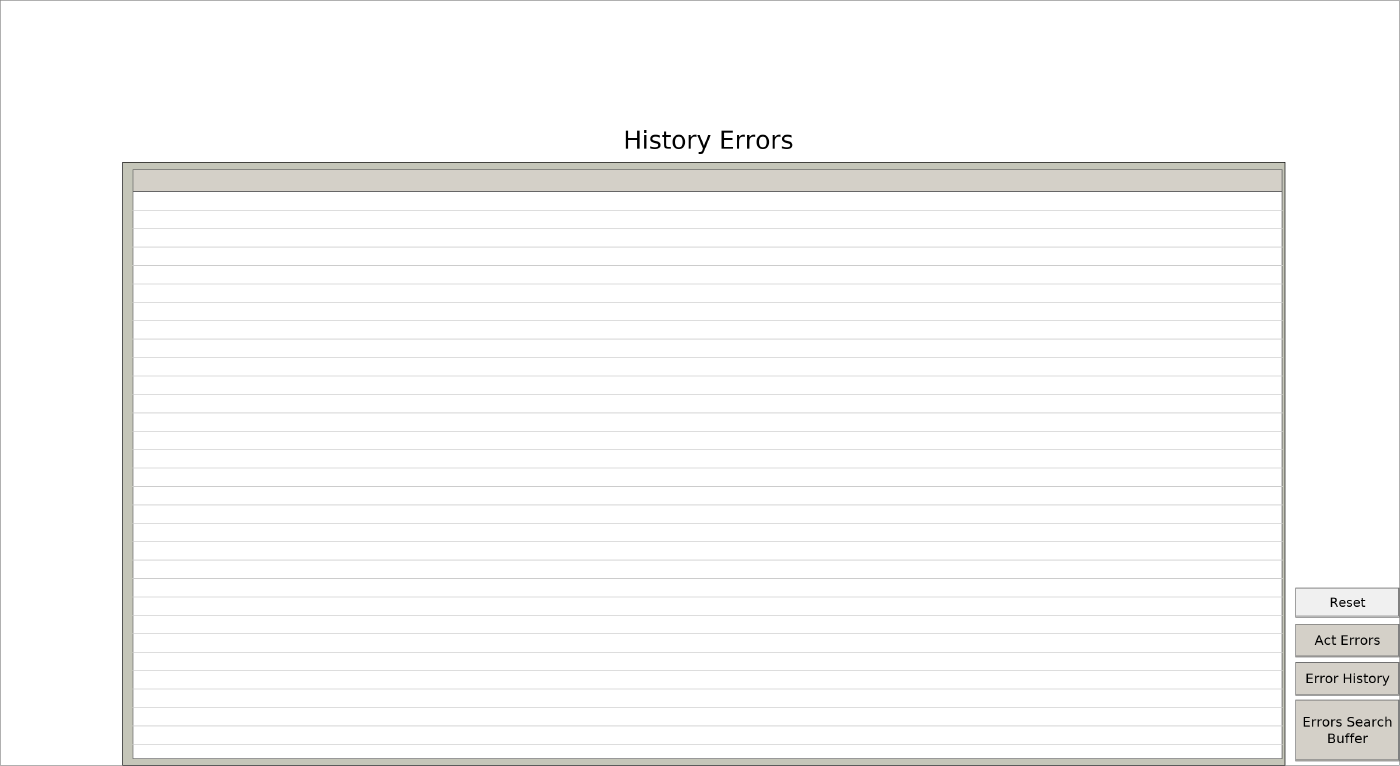
VISUALIZATION ERROR_HISTORY  // 1900x1040
    Group (1758,798 142x235)
        Button (0,0 142x40), "Reset", pressed state: prg_Messages.ResetErrors
            toggle prg_Messages.ResetErrors
        Button (0,101 142x45), "Error History"
            OnMouseClick: change screen: ERROR_HISTORY
        Button (0,152 142x83), "Errors Search Buffer"
            OnMouseClick: change screen: ERROR_BUFFER
        Button (0,49 142x45), "Act Errors"
            OnMouseClick: change screen: ERRORS_OPER
    Rectangle (166,220 1578x820)
    Rectangle (841,165 241x50), "History Errors"
    Table (180,230 1560x800), data array: Buffer_Act_History
        p3854506369: Buffer_Act_History[INDEX].sDateTime
        p1892666644: Buffer_Act_History[INDEX].sErrID
        p338671338: Buffer_Act_History[INDEX].sLevel
        p2170511999: Buffer_Act_History[INDEX].sModuleDescription
        p3723444502: Buffer_Act_History[INDEX].sErrorMessage
        p4092479075: Module Description
        p2237128397: Error Message
END_VISUALIZATION

(* stored: Version 1.1.0.1, ProductVersion 3.1.4024.13
   Visu ERROR_HISTORY: Id {9c6edd7a-4ebf-4f41-bf25-672af31ad049} *)
